ABB RobotStudio station: project1.rspag

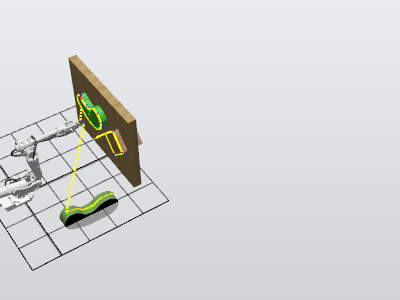
--- station ---
Station Projekt_pierwszy (saved by RobotStudio 24.3.10958.1)
Controller Controller1
  mechanical unit ROB_1: IRB6650S_125_350_MH3_03, 6 joints, base frame (0, 0, 0) mm
Layout (positions relative to the parent item):
  - IRB6650S_125_350_MH3_03 [mechanism, from %ABB.RobotStudio.Models.IRB6650S%\IRB6650S_125_350_MH3_03.rslib] at (0, 0, 0) mm; joint values [0, 0, 0, 0, 0.5236, 0] (rad or m)
  - Group_2 [graphiccomponentgroup] at (2365.21, 0, 2010) mm, rotated rx 180 ry 60 rz 180 deg
    - Part_6 [part] at (-29.38, 0.12, 253.59) mm, rotated rx -45 ry 0 rz 90 deg, size 40 x 39.7 x 50 mm
    - Part_2 [part], size 200 x 198.9 x 40 mm
    - Part_4 [part] at (0, 0, 33.32) mm, size 40 x 40 x 200 mm
    - Part_5 [part] at (5.57, 0.1, 219.05) mm, rotated rx -45 ry 0 rz 90 deg, size 40 x 39.7 x 50 mm
  - Part_8 [part] at (3927.17, -1627.08, 1612.93) mm, rotated rx -90 ry -46.19 rz 90 deg, size 780 x 780 x 780 mm
  - Part_11 [part] at (3514.72, 422.88, 1806.86) mm, rotated rx 0 ry -90 rz 0 deg, size 886.3 x 1638.1 x 400 mm
  - Part_12 [part] at (3341.47, -1836.92, 0) mm, size 300 x 4000 x 3000 mm
  - Part_14 [part] at (1609.3, -1676.33, 0) mm, rotated rx 0 ry -90 rz 90 deg, size 875.9 x 1971.5 x 400 mm
Attachment: Group_2 is attached to IRB6650S_125_350_MH3_03 / Link6
Attachment: Block is attached to Part_8
Attachment: OnTheWall is attached to Part_11
Attachment: OnTheFloor is attached to Part_14
Collision set CollisionSet_1: IRB6650S_125_350_MH3_03, Group_2 against Part_8, Part_11, Part_12, Part_14, near miss 0 m
Targets, tools, work objects and paths stored in the station and not in the controller backup, written as RAPID:
! task T_ROB1
MODULE Module1
  CONST robtarget Target_10:=[[-0.000827752,779.999086422,0],[0,0.919852246,0.39226502,0],[-1,1,0,0],[9E+09,9E+09,9E+09,9E+09,9E+09,9E+09]];
  CONST robtarget Target_20:=[[779.99895192,780.0007937,0],[0,0.919852246,0.39226502,0],[-1,0,1,0],[9E+09,9E+09,9E+09,9E+09,9E+09,9E+09]];
  CONST robtarget Target_30:=[[779.99996694,0.000292377,0],[0,0.919852246,0.39226502,0],[-1,1,0,0],[9E+09,9E+09,9E+09,9E+09,9E+09,9E+09]];
  CONST robtarget Target_40:=[[0.000157874,-0.000000992,0],[0,0.919852246,0.39226502,0],[-1,1,0,0],[9E+09,9E+09,9E+09,9E+09,9E+09,9E+09]];
  CONST robtarget Target_60:=[[97.52923891,513.47613776,472.353802441],[0.516842609,-0.228370254,-0.418040767,0.711310524],[0,-2,-2,0],[9E+09,9E+09,9E+09,9E+09,9E+09,9E+09]];
  CONST robtarget Target_70:=[[47.693410332,634.01244556,482.431760765],[0.468024692,-0.25586516,-0.40180104,0.744339863],[0,-2,-2,0],[9E+09,9E+09,9E+09,9E+09,9E+09,9E+09]];
  CONST robtarget Target_80:=[[-20.890984187,743.760617829,459.439970741],[0.286847755,-0.340392124,-0.333233038,0.831148187],[0,-1,-2,0],[9E+09,9E+09,9E+09,9E+09,9E+09,9E+09]];
  CONST robtarget Target_90:=[[-146.663361904,808.37254164,327.546222241],[0.107505923,0.452189201,0.149786457,-0.872657677],[0,-1,-1,0],[9E+09,9E+09,9E+09,9E+09,9E+09,9E+09]];
  CONST robtarget Target_100:=[[-224.111368116,727.420855901,167.045312064],[0.50239854,0.469823197,-0.078595292,-0.721584819],[0,-1,-1,0],[9E+09,9E+09,9E+09,9E+09,9E+09,9E+09]];
  CONST robtarget Target_110:=[[-223.295805372,702.314491867,151.689459989],[0.585937236,0.456877948,-0.134809481,-0.655565786],[0,-1,-1,0],[9E+09,9E+09,9E+09,9E+09,9E+09,9E+09]];
  CONST robtarget Target_120:=[[-218.228254946,674.762055216,140.620669922],[0.645395079,0.442055526,-0.177476668,-0.597121543],[0,-1,0,0],[9E+09,9E+09,9E+09,9E+09,9E+09,9E+09]];
  CONST robtarget Target_130:=[[-198.761735053,614.153311713,127.802364835],[0.706460488,0.420151951,-0.224462455,-0.523452503],[0,-1,0,0],[9E+09,9E+09,9E+09,9E+09,9E+09,9E+09]];
  CONST robtarget Target_140:=[[-146.474827093,483.760777463,114.649478077],[0.701996867,0.422040012,-0.22089202,-0.529423595],[0,-1,0,0],[9E+09,9E+09,9E+09,9E+09,9E+09,9E+09]];
  CONST robtarget Target_150:=[[-109.646937222,303.675248066,47.439097823],[0.560820927,0.461632859,-0.117499615,-0.677177105],[0,-2,0,0],[9E+09,9E+09,9E+09,9E+09,9E+09,9E+09]];
  CONST robtarget Target_160:=[[-107.793488854,187.403858868,-26.342238963],[0.510837181,0.468867891,-0.084106817,-0.715635605],[0,-2,0,0],[9E+09,9E+09,9E+09,9E+09,9E+09,9E+09]];
  CONST robtarget Target_170:=[[-138.891493582,79.32265082,-140.41642514],[0.269391498,0.472266979,0.062249149,-0.836969035],[0,-1,-1,0],[9E+09,9E+09,9E+09,9E+09,9E+09,9E+09]];
  CONST robtarget Target_180:=[[-152.912822957,69.365795516,-166.388321438],[0.20254836,0.465887138,0.099298693,-0.855606864],[0,-1,-1,0],[9E+09,9E+09,9E+09,9E+09,9E+09,9E+09]];
  CONST robtarget Target_190:=[[-223.327609288,50.137148866,-276.61036853],[0.155719516,0.45979773,0.12448736,-0.865355636],[0,-1,-2,0],[9E+09,9E+09,9E+09,9E+09,9E+09,9E+09]];
  CONST robtarget Target_200:=[[-280.283568082,3.692528594,-386.049888704],[0.349160793,0.476075179,0.016232056,-0.806954574],[0,-1,-2,0],[9E+09,9E+09,9E+09,9E+09,9E+09,9E+09]];
  CONST robtarget Target_210:=[[-281.299044454,-264.466887573,-563.545665018],[0.670820922,0.433895425,-0.196585392,-0.56840851],[-1,0,-2,0],[9E+09,9E+09,9E+09,9E+09,9E+09,9E+09]];
  CONST robtarget Target_220:=[[-121.666754724,-543.973583739,-525.833613631],[0.852918634,0.302413765,-0.368044795,-0.213585458],[-1,1,-2,0],[9E+09,9E+09,9E+09,9E+09,9E+09,9E+09]];
  CONST robtarget Target_230:=[[5.16591795,-609.639771566,-393.162576014],[0.878718575,0.18879548,-0.437341197,0.030701942],[-1,1,-2,0],[9E+09,9E+09,9E+09,9E+09,9E+09,9E+09]];
  CONST robtarget Target_240:=[[123.106834385,-598.840339146,-222.604023777],[0.861772285,0.114479191,-0.462391145,0.174463386],[-1,1,-2,0],[9E+09,9E+09,9E+09,9E+09,9E+09,9E+09]];
  CONST robtarget Target_250:=[[231.092359404,-498.477813785,-7.031638074],[0.80043741,0.007527124,-0.476292345,0.36385285],[0,2,-2,0],[9E+09,9E+09,9E+09,9E+09,9E+09,9E+09]];
  CONST robtarget Target_260:=[[270.989744042,-312.298064132,170.522384521],[0.721112189,-0.079036944,-0.4697491,0.50307669],[0,2,-2,0],[9E+09,9E+09,9E+09,9E+09,9E+09,9E+09]];
  CONST robtarget Target_270:=[[269.709101767,-87.792063109,316.170473108],[0.673093489,-0.120843257,-0.460768883,0.565715564],[0,2,-2,0],[9E+09,9E+09,9E+09,9E+09,9E+09,9E+09]];
  CONST robtarget Target_280:=[[230.753641151,148.642651228,417.43401774],[0.584590773,-0.185950859,-0.438558245,0.656766756],[0,2,-2,0],[9E+09,9E+09,9E+09,9E+09,9E+09,9E+09]];
  CONST robtarget Target_290:=[[192.577241102,269.625105887,443.965001348],[0.535450812,-0.217248458,-0.423927073,0.697410476],[0,2,-2,0],[9E+09,9E+09,9E+09,9E+09,9E+09,9E+09]];
  CONST robtarget Target_300:=[[97.52923891,513.47613776,472.353802441],[0.516842609,-0.228370254,-0.418040767,0.711310524],[0,2,-2,0],[9E+09,9E+09,9E+09,9E+09,9E+09,9E+09]];
  CONST robtarget Target_310:=[[1798.032513692,-2268.256416295,1872.178062751],[0.312844431,0.657136635,0.572149215,-0.378080787],[-1,0,-1,0],[9E+09,9E+09,9E+09,9E+09,9E+09,9E+09]];
  CONST robtarget Target_320:=[[292.788251262,613.280476419,494.594671725],[0.001140751,-0.65191797,0.758137413,0.015143383],[0,0,0,0],[9E+09,9E+09,9E+09,9E+09,9E+09,9E+09]];
  CONST robtarget Target_330:=[[269.970225826,508.288710879,463.679735882],[0.001140751,-0.65191797,0.758137413,0.015143383],[0,0,0,0],[9E+09,9E+09,9E+09,9E+09,9E+09,9E+09]];
  CONST robtarget Target_340:=[[273.750189703,419.311313125,416.455695414],[0.001140751,-0.65191797,0.758137413,0.015143383],[0,0,0,0],[9E+09,9E+09,9E+09,9E+09,9E+09,9E+09]];
  CONST robtarget Target_350:=[[282.270148249,313.714871939,326.05974192],[0.001140751,-0.65191797,0.758137413,0.015143383],[0,0,0,0],[9E+09,9E+09,9E+09,9E+09,9E+09,9E+09]];
  CONST robtarget Target_360:=[[274.725620007,225.530944313,212.003639837],[0.001140751,-0.65191797,0.758137413,0.015143383],[0,0,0,0],[9E+09,9E+09,9E+09,9E+09,9E+09,9E+09]];
  CONST robtarget Target_370:=[[244.279320632,117.275094291,165.415147168],[0.001140751,-0.65191797,0.758137413,0.015143383],[0,0,0,0],[9E+09,9E+09,9E+09,9E+09,9E+09,9E+09]];
  CONST robtarget Target_380:=[[211.52196329,-57.049702716,155.377572811],[0.001140751,-0.65191797,0.758137413,0.015143383],[0,0,0,0],[9E+09,9E+09,9E+09,9E+09,9E+09,9E+09]];
  CONST robtarget Target_390:=[[155.521214817,-213.936273695,219.64189925],[0.001140751,-0.65191797,0.758137413,0.015143383],[0,0,0,0],[9E+09,9E+09,9E+09,9E+09,9E+09,9E+09]];
  CONST robtarget Target_400:=[[140.800461683,-345.059788734,299.383517542],[0.001140751,-0.65191797,0.758137413,0.015143383],[0,0,0,0],[9E+09,9E+09,9E+09,9E+09,9E+09,9E+09]];
  CONST robtarget Target_410:=[[111.511458878,-570.494709389,355.980499044],[0.001140751,-0.65191797,0.758137413,0.015143383],[0,0,0,0],[9E+09,9E+09,9E+09,9E+09,9E+09,9E+09]];
  CONST robtarget Target_420:=[[88.423436997,-756.468950878,326.500378707],[0.001140751,-0.65191797,0.758137413,0.015143383],[0,0,0,0],[9E+09,9E+09,9E+09,9E+09,9E+09,9E+09]];
  CONST robtarget Target_430:=[[101.349410687,-930.117750769,242.553332311],[0.001140751,-0.65191797,0.758137413,0.015143383],[0,0,0,0],[9E+09,9E+09,9E+09,9E+09,9E+09,9E+09]];
  CONST robtarget Target_440:=[[314.516037972,757.824115529,492.465304984],[0.001140751,-0.65191797,0.758137413,0.015143383],[0,0,0,0],[9E+09,9E+09,9E+09,9E+09,9E+09,9E+09]];
  CONST robtarget Target_310_2:=[[507.651484902,256.805488593,537.163983175],[0.945065405,0.281129847,-0.160261192,-0.046192416],[-1,0,-1,0],[9E+09,9E+09,9E+09,9E+09,9E+09,9E+09]];
  CONST robtarget Target_310_2_2:=[[1931.936016853,-1385.894468812,1891.347424043],[0.312844431,0.657136635,0.572149215,-0.378080787],[-1,0,-1,0],[9E+09,9E+09,9E+09,9E+09,9E+09,9E+09]];
  CONST robtarget Target_10_2:=[[-0.000827752,779.999086422,421.130610934],[0,0.919852246,0.39226502,0],[-1,1,0,0],[9E+09,9E+09,9E+09,9E+09,9E+09,9E+09]];
  PROC Path_10()
    MoveL Target_10,v1000,fine,swieczka\WObj:=Block;
    MoveL Target_20,v500,fine,swieczka\WObj:=Block;
    MoveL Target_30,v500,fine,swieczka\WObj:=Block;
    MoveL Target_40,v500,fine,swieczka\WObj:=Block;
    MoveL Target_10,v500,fine,swieczka\WObj:=Block;
    MoveL Target_10_2,v1000,z0,swieczka\WObj:=Block;
  ENDPROC
  PROC Path_20()
    MoveL Target_60,v1000,z10,swieczka\WObj:=OnTheWall;
    MoveC Target_70,Target_80,v800,z10,swieczka\WObj:=OnTheWall;
    MoveC Target_90,Target_100,v800,z10,swieczka\WObj:=OnTheWall;
    MoveL Target_110,v800,z10,swieczka\WObj:=OnTheWall;
    MoveL Target_120,v800,z10,swieczka\WObj:=OnTheWall;
    MoveL Target_130,v800,z10,swieczka\WObj:=OnTheWall;
    MoveC Target_140,Target_150,v800,z10,swieczka\WObj:=OnTheWall;
    MoveC Target_160,Target_170,v800,z10,swieczka\WObj:=OnTheWall;
    MoveL Target_180,v800,z10,swieczka\WObj:=OnTheWall;
    MoveC Target_190,Target_200,v800,z10,swieczka\WObj:=OnTheWall;
    MoveC Target_210,Target_220,v800,z10,swieczka\WObj:=OnTheWall;
    MoveC Target_230,Target_240,v800,z10,swieczka\WObj:=OnTheWall;
    MoveC Target_250,Target_260,v800,z10,swieczka\WObj:=OnTheWall;
    MoveC Target_270,Target_280,v800,z10,swieczka\WObj:=OnTheWall;
    MoveL Target_290,v800,z10,swieczka\WObj:=OnTheWall;
    MoveL Target_300,v800,z10,swieczka\WObj:=OnTheWall;
    MoveJ Target_310_2,v1000,z50,swieczka\WObj:=OnTheWall;
  ENDPROC
  PROC Path_30()
    MoveJ Target_430,v1000,z10,swieczka\WObj:=OnTheFloor;
    MoveL Target_420,v400,z10,swieczka\WObj:=OnTheFloor;
    MoveL Target_410,v400,z10,swieczka\WObj:=OnTheFloor;
    MoveL Target_400,v400,z10,swieczka\WObj:=OnTheFloor;
    MoveL Target_390,v400,z10,swieczka\WObj:=OnTheFloor;
    MoveL Target_380,v400,z10,swieczka\WObj:=OnTheFloor;
    MoveL Target_370,v400,z10,swieczka\WObj:=OnTheFloor;
    MoveL Target_360,v400,z10,swieczka\WObj:=OnTheFloor;
    MoveL Target_350,v400,z10,swieczka\WObj:=OnTheFloor;
    MoveL Target_340,v400,z10,swieczka\WObj:=OnTheFloor;
    MoveL Target_330,v400,z10,swieczka\WObj:=OnTheFloor;
    MoveL Target_320,v400,z10,swieczka\WObj:=OnTheFloor;
    MoveL Target_440,v400,z50,swieczka\WObj:=OnTheFloor;
    WaitTime 0.1;
    MoveJ Target_310_2_2,v1000,z100,swieczka\WObj:=OnTheFloor;
  ENDPROC
ENDMODULE

! task T_ROB1
MODULE CalibData
  TASK PERS wobjdata Block:=[FALSE,TRUE,"",[[3147.174649931,-1064.191574427,1072.966259915],[0.650433761,0.277373256,-0.650433761,-0.277373256]],[[0,0,0],[1,0,0,0]]];
  TASK PERS wobjdata OnTheWall:=[FALSE,TRUE,"",[[3114.719771138,430.591427426,1800.955],[0.333742439,-0.100561118,0.898581245,0.266561797]],[[0,0,0],[1,0,0,0]]];
  TASK PERS wobjdata OnTheFloor:=[FALSE,TRUE,"",[[1608.579096564,-2076.33,-37.839],[0.65191797,-0.001140751,-0.015143383,0.758137413]],[[0,0,0],[1,0,0,0]]];
ENDMODULE


--- Controller Data/Controller1/RAPID/TASK1/PROGMOD/Module1.mod ---
MODULE Module1
	TASK PERS tooldata swieczka:=[TRUE,[[-64.6298,0.0716233,289.296],[1,0,0,0]],[1,[0,0,0],[1,0,0,0],0,0,0]];
    !***********************************************************
    !
    ! Module:  Module1
    !
    ! Description:
    !   <Insert description here>
    !
    ! Author: Mirgi
    !
    ! Version: 1.0
    !
    !***********************************************************


    !***********************************************************
    !
    ! Procedure main
    !
    !   This is the entry point of your program
    !
    !***********************************************************
    PROC main()
        !Add your code here
    ENDPROC
ENDMODULE
